FUNCTION_BLOCK DrillingSequence (* Composite Function Block Type *)
  (* Standard: 61499-2 *)
  (* Version 0.0, 7/2/2026, template *)
  PACKAGE Main;
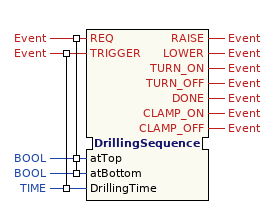
  EVENT_INPUT
    REQ WITH atTop, atBottom; (* Normal Execution Request *)
    TRIGGER WITH DrillingTime;
  END_EVENT
  EVENT_OUTPUT
    RAISE; (* Initialization Confirm *)
    LOWER; (* Execution Confirmation *)
    TURN_ON;
    TURN_OFF;
    DONE;
    CLAMP_ON;
    CLAMP_OFF;
  END_EVENT
  VAR_INPUT
    atTop : BOOL; (* Input event qualifier *)
    atBottom : BOOL;
    DrillingTime : TIME;
  END_VAR
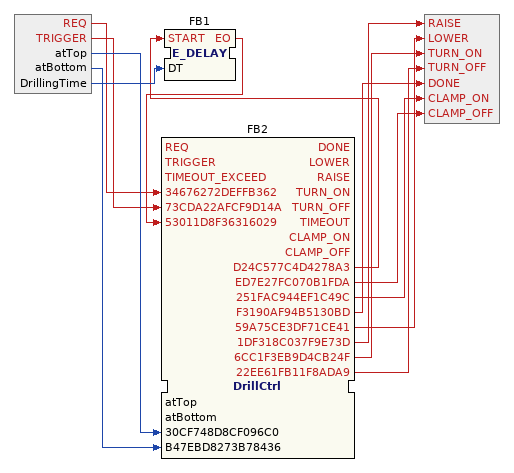
  FBS
    FB1 : E_DELAY;
    FB2 : DrillCtrl;
  END_FBS
  EVENT_CONNECTIONS
    REQ TO FB2.34676272DEFFB362;
    TRIGGER TO FB2.73CDA22AFCF9D14A;
    FB1.EO TO FB2.53011D8F36316029;
    FB2.D24C577C4D4278A3 TO FB1.START;
    FB2.ED7E27FC070B1FDA TO CLAMP_OFF;
    FB2.251FAC944EF1C49C TO CLAMP_ON;
    FB2.F3190AF94B5130BD TO DONE;
    FB2.59A75CE3DF71CE41 TO LOWER;
    FB2.1DF318C037F9E73D TO RAISE;
    FB2.6CC1F3EB9D4CB24F TO TURN_ON;
    FB2.22EE61FB11F8ADA9 TO TURN_OFF;
  END_CONNECTIONS
  DATA_CONNECTIONS
    DrillingTime TO FB1.DT;
    atTop TO FB2.30CF748D8CF096C0;
    atBottom TO FB2.B47EBD8273B78436;
  END_CONNECTIONS
END_FUNCTION_BLOCK
